// TIA Portal V20 export
DATA_BLOCK "Global_Signal"   // DB41
{ S7_Optimized_Access := 'FALSE' }
   VAR
      "M_Grundstellung_POS3.0" : Bool := TRUE;
   END_VAR
BEGIN
END_DATA_BLOCK
